(* IEC 61131-3 sources: kns-port-domestic/upstream/plc-process-lib/src/POUs/Util/F_LTimeToSec, 1 file *)

(* ---- F_LTimeToSec.decl.st ---- *)
// Назначение: длительность LTIME (нс) в секундах LREAL. LTIME без знака: отрицательных
//             значений не бывает, разность отметок вызывающий считает только при a >= b.
// Автор:      kr0nsch
// Версия:     0.1.0
// Документ:   docs/fb/Functions.md
FUNCTION F_LTimeToSec : LREAL
VAR_INPUT
    ltIn : LTIME;   // длительность или разность монотонных отметок
END_VAR
